// This function has been automatically generated from the project information.
{attribute 'signature_flag' := '1073741824'}
{attribute 'TcGenerated'}
{attribute 'no-analysis'}
FUNCTION F_GetVersion : ST_LibVersion
VAR_INPUT
	
END_VAR

F_GetVersion.iMajor := 1;
F_GetVersion.iMinor := 2;
F_GetVersion.iBuild := 0;
F_GetVersion.iRevision := 0;
F_GetVersion.sVersion := '1.2.0';
F_GetVersion.nFlags := 1;

END_FUNCTION

(* stored: Version 1.1.0.1
   POU F_GetVersion: Id {6cec820c-0b6c-017e-278d-f0a5ea844896}, SpecialFunc None *)
